(* IEC 61131-3 sources: trust-platform/examples/OSCAT/ventilation_filter/non-oop/src, 3 files *)

(* ---- Configuration.st ---- *)
CONFIGURATION VentilationFilterClassicConfiguration
RESOURCE Cpu0 ON PLC
    TASK MainTask (INTERVAL := T#100ms, PRIORITY := 1);
    PROGRAM Main WITH MainTask : Main;
END_RESOURCE
END_CONFIGURATION

(* ---- Main.st ---- *)
PROGRAM Main
VAR
    IntakeFilter : FT_PT1;
    ExhaustFilter : FT_PT1;
    RawAirflow : REAL := REAL#10.0;
    IntakeAirflow : REAL;
    ExhaustAirflow : REAL;
END_VAR

IntakeFilter(in := RawAirflow, T := T#1s, K := REAL#1.0);
ExhaustFilter(in := RawAirflow, T := T#1s, K := REAL#2.0);
IntakeAirflow := IntakeFilter.out;
ExhaustAirflow := ExhaustFilter.out;
END_PROGRAM

(* ---- Tests.st ---- *)
TEST_PROGRAM VentilationFilterClassicKeepsTwoFilterInstancesIndependent
VAR
    IntakeFilter : FT_PT1;
    ExhaustFilter : FT_PT1;
END_VAR

IntakeFilter(in := REAL#10.0, T := T#1s, K := REAL#1.0);
ExhaustFilter(in := REAL#10.0, T := T#1s, K := REAL#2.0);

ASSERT_NEAR(EXPECTED := REAL#10.0, ACTUAL := IntakeFilter.out, DELTA := REAL#0.001);
ASSERT_NEAR(EXPECTED := REAL#20.0, ACTUAL := ExhaustFilter.out, DELTA := REAL#0.001);
END_TEST_PROGRAM
